Fanuc KAREL source: KT00761.KL

PROGRAM KT00761
%NOLOCKGROUP
VAR
  I1: INTEGER
  I2: INTEGER
  OUT: REAL
BEGIN
  I1 = 2
  I2 = 3
  I1 = 2
  I2 = 3
  OUT = ACOS(I1)
END KT00761
